(* Simple NOT Gate Operation *)

PROGRAM main
  VAR
    Input AT %IX0.6 : BOOL;
    Output AT %QX0.3 : BOOL;
  END_VAR

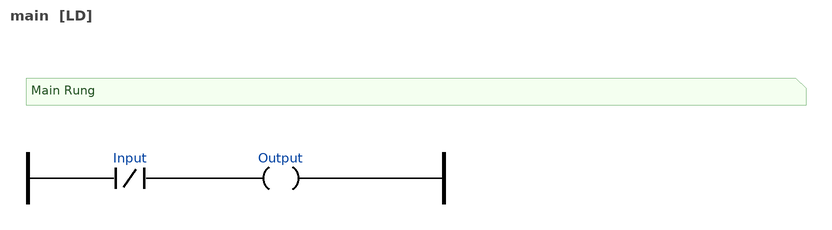
(* LD diagram, written out as Structured Text *)
(* Main Rung *)
Output := NOT Input;
END_PROGRAM
